// TIA Portal V20 export
Screen "11_SubMenus_Type"  100x768
  ScreenItem "txtOverview_1" at -1,554 size 100x41  Type=HmiTextBox
  ScreenItem "txtOverview_2" at -1,490 size 100x49  Type=HmiTextBox
  ScreenItem "txtOverview_3" at 394,557 size 100x41  Type=HmiTextBox
  ScreenItem "txtOverview_4" at -1,441 size 100x43  Type=HmiTextBox
  ScreenItem "txtOverview_5" at -1,393 size 100x42  Type=HmiTextBox
  ScreenItem "txtOverview_6" at -1,339 size 100x52  Type=HmiTextBox
  ScreenItem "txtOverview_7" at -1,283 size 100x52  Type=HmiTextBox
  ScreenItem "txtOverview_8" at -1,224 size 100x52  Type=HmiTextBox
  ScreenItem "txtOverview_9" at -1,167 size 100x52  Type=HmiTextBox
  ScreenItem "txtOverview_10" at -1,108 size 100x52  Type=HmiTextBox
  ScreenItem "txtOverview_11" at -1,53 size 100x52  Type=HmiTextBox
  ScreenItem "txtOverview_12" at -1,-7 size 100x52  Type=HmiTextBox
  ScreenItem "线_1" at -1,391 size 97x0  Type=HmiLine
  ScreenItem "txtOverview_13" at -1,546 size 100x49  Type=HmiTextBox
  ScreenItem "txtOverview_15" at -1,711 size 100x49  Type=HmiTextBox
  ScreenItem "txtOverview_16" at -1,655 size 100x49  Type=HmiTextBox
  ScreenItem "txtOverview_14" at -1,607 size 100x41  Type=HmiTextBox
  ScreenItem "txtOverview_17" at -1,599 size 100x49  Type=HmiTextBox
